(* Logix 5000 project; controller DSFW_Budzar vendor 1 type 14 code 154 rev 32.13; software revision 32.03; part 2 of 5 *)
(* tags used below, declared in another part *)
   ACKNOWLEDGE_ALARMS : BOOL;
   Active_Setpoint : REAL;
   ALARMS : DINT[5];
   ALWAYS_OFF : BOOL;
   Batch_High_High_Temp_Delay : TIMER;
   Batch_High_High_Temp_Setpoint : REAL;
   Batch_Jacket_DT_Temp_Delay : TIMER;
   Batch_Low_Low_Temp_Delay : TIMER;
   Batch_Low_Low_Temp_Setpoint : REAL;
   Batch_Mode_Enable : BOOL;
   C1_Low_Oil_Timer : TIMER;
   C1_MP_Timer : TIMER;
   C1_Run_Proof_Timer : TIMER;
   C_101_AUX : ALIAS FOR Local:1:I.Data.8;
   Comp_Start_Purge_Relay : BOOL;
   Compressor_R404A_Superheat : REAL;
   Condenser_Water_Inlet_Temp_Limit : REAL;
   Condenser_Water_Inlet_Temp_TMR : TIMER;
   CR_002 : ALIAS FOR Local:1:I.Data.0;   // Emergency Stop Safety Relay Status
   CR_01 : ALIAS FOR Local:1:I.Data.15;   // Glycol Tank Low Level Alarm Relay Dry Contact
   CR_108 : ALIAS FOR Local:1:O.Data.0;   // Process Pump Motor Relay (Energizes Contactor M-101)
   CR_109 : ALIAS FOR Local:1:O.Data.5;   // Compressor Motor Relay (Energizes Contactor C-101)
   DCS_Comm_TMR : TIMER;
   DCS_Heartbeat_Returned : DINT;
   DCS_Heartbeat_Returned_Last : DINT;
   EEV_Manual_Relief_Delay : TIMER;   // Oil Management, Delay until Flush begins
   EEV_Manual_Relief_Timer : TIMER;   // Oil Management, Duration of Flush
   FIC_101_Run_PID : BOOL;
   HMI_Batch_Hi_Hi_Temp_Delay : DINT;
   HMI_Batch_Jacket_DT_Temp_Delay : DINT;
   HMI_Batch_Low_Low_Temp_Delay : DINT;
   HMI_Condenser_Water_Inlet_Temp_Delay : DINT;
   HMI_EEV_Manual_Relief_Delay : REAL;   // Oil Management, Delay to start relief entered in minutes.
   HMI_EEV_Manual_Relief_Timer : REAL;   // Oil Management, Relief Duration entered in seconds
   HMI_Jacket_Hi_Hi_Temp_Delay : DINT;
   HMI_Jacket_Hi_Temp_Delay : REAL;
   HMI_Jacket_Low_Low_Temp_Delay : DINT;
   HMI_Jacket_Low_Temp_Delay : REAL;
   HMI_Low_Pump_Suction_Pressure_Delay : REAL;
   HMI_PCV_101_Flush_Time : DINT;
   HMI_R507A_High_Superheat_Timer : DINT;
   HMI_R507A_Low_Pressure_Delay : DINT;
   HMI_R507A_Low_Superheat_Timer : DINT;
   HMI_Remote_State_1 : BOOL;
   HMI_Remote_State_2 : BOOL;
   HMI_Return_Trend_Limits : REAL[2];
   HMI_SP_Trend_Limits : REAL[2];
   HMI_Supply_Trend_Limits : REAL[2];
   HMI_Trend_Data : REAL[3];
   HMI_Valve_Flush_SP : REAL;
   Jacket_Batch_Delta_T : REAL;
   Jacket_Batch_High_Delta_T_Setpoint : REAL;
   Jacket_High_High_Temp_Delay : TIMER;
   Jacket_High_High_Temp_Setpoint : REAL;
   Jacket_High_Temp_Delay : TIMER;
   Jacket_High_Temp_Setpoint : REAL;
   Jacket_Low_Low_Temp_Delay : TIMER;
   Jacket_Low_Low_Temp_Setpoint : REAL;
   Jacket_Low_Temp_Delay : TIMER;
   Jacket_Low_Temp_Setpoint : REAL;
   Low_Pump_Suction_Pressure_Delay : TIMER;
   Low_Pump_Suction_Pressure_Setpoint : REAL;
   M_101_AUX : ALIAS FOR Local:1:I.Data.3;
   Oil_Purge_Fail : BOOL;   // Oil Management, This coil will energize after configured purge retries fail
   Oil_Purge_Retires_Enable : BOOL;
   OMB_101 : ALIAS FOR Local:1:I.Data.12;
   PCV_101_Flush_Timer : TIMER;   // PCV-101 Condenser Hot Water Flush Timer
   PM_101 : ALIAS FOR Local:1:I.Data.1;
   PM_101_StartupTMR : TIMER;   // PM-101 Phase Monitor Startup Delay Alarm Timer
   Process_Pump_Diff_Pressure : REAL;
   PT_101 : BL_Analog_Input;   // Process Supply Pressure
   PT_102 : BL_Analog_Input;   // R404A Compressor Suction Pressure
   PT_103 : BL_Analog_Input;   // R404A Compressor Discharge Pressure
   PT_105 : BL_Analog_Input;   // Condenser Chilled Glycol Return Pressure
   PT_107 : BL_Analog_Input;   // Process Pump Suction Pressure
   Pump_1_Low_Press_Delay : TIMER;
   Pump_High_Pressure_Alarm_Setpoint : REAL;
   Pump_Low_Pressure_Alarm_Setpoint : REAL;
   Pump_RP_ALM_TMR : TIMER;
   R404A_High_Pressure_Setpoint : REAL;
   R404A_High_SH_Setpoint : REAL;
   R404A_High_Superheat_Timer : TIMER;
   R404A_Low_Pressure_Delay : TIMER;
   R404A_Low_Pressure_Setpoint : REAL;
   R404A_Low_SH_Setpoint : REAL;
   R404A_Low_Superheat_Timer : TIMER;
   Ramp_Soak_Current_HMI : DINT;
   Ramp_Soak_Segments_HMI : DINT;
   Ramp_Soak_Segments_HMI_Set : REAL;
   Remote_System_Start : BOOL;   // Remote Start/Stop 0=Stop 1=Start
   Remote_Temp_Setpoint : REAL;   // Remote Temperature Setpoint
   RX_RMPS : RAMP_SOAK;
   Slot_2_Status : DINT;
   Slot_3_Status : DINT;
   Slot_4_Status : DINT;
   Slot_5_Status : DINT;
   Slot_6_Status : DINT;
   Slot_7_Status : DINT;
   Slot_8_Status : DINT;
   Slot_9_Status : DINT;
   Start_Up_Delay : TIMER;
   System_Mode : BOOL;   // 0 = Local Control 1 = Remote Control
   TE_101 : BL_Analog_Input;   // Process Supply Temperature
   TE_102 : BL_Analog_Input;   // Process Return Temperature
   TE_108 : BL_Analog_Input;   // CONDENSER CHILLED GLYCOL INLET TEMPERATURE SENSOR
   Temperature_Setpoint_Max : REAL;   // Maximum Operating Temperature Setpoint (Deg C)
   Temperature_Setpoint_Min : REAL;   // Minimum Operating Temperature Setpoint (Deg C)
   TSH_101 : ALIAS FOR Local:1:I.Data.4;
   Valve_delay_count : REAL;
   Valve_Flush_SP : REAL;
   VESSEL_TEMPERATURE : BL_Analog_Input;   // End User Reactor Temperature
(* A_MainProgram, continued *)

ROUTINE General_Process_Alarms   (* ladder *)
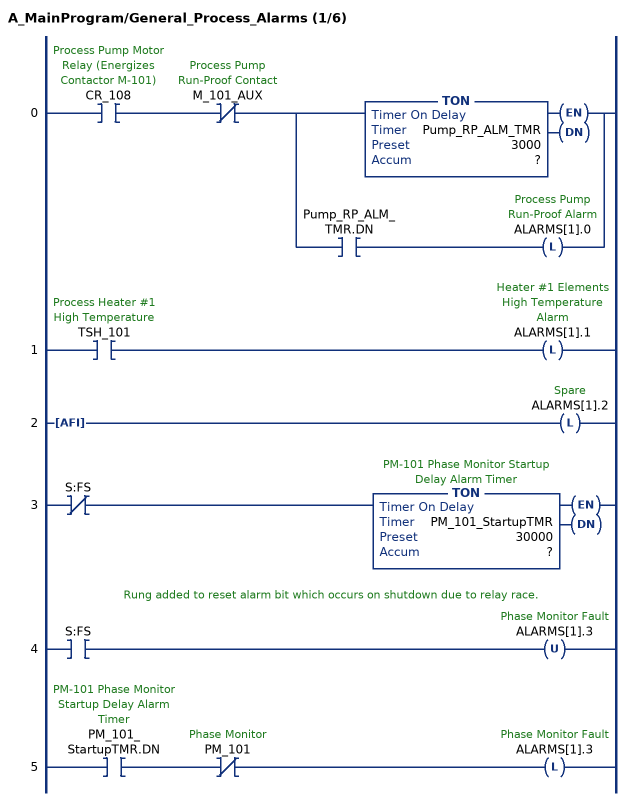
   0: XIC(CR_108)XIO(M_101_AUX)[TON(Pump_RP_ALM_TMR,?,?) ,XIC(Pump_RP_ALM_TMR.DN) OTL(ALARMS[1].0) ];
   1: XIC(TSH_101)OTL(ALARMS[1].1);
   2: AFI()OTL(ALARMS[1].2);
   3: XIO(S:FS)TON(PM_101_StartupTMR,?,?);
   // Rung added to reset alarm bit which occurs on shutdown due to relay race.
   4: XIC(S:FS)OTU(ALARMS[1].3);
   5: XIC(PM_101_StartupTMR.DN)XIO(PM_101)OTL(ALARMS[1].3);
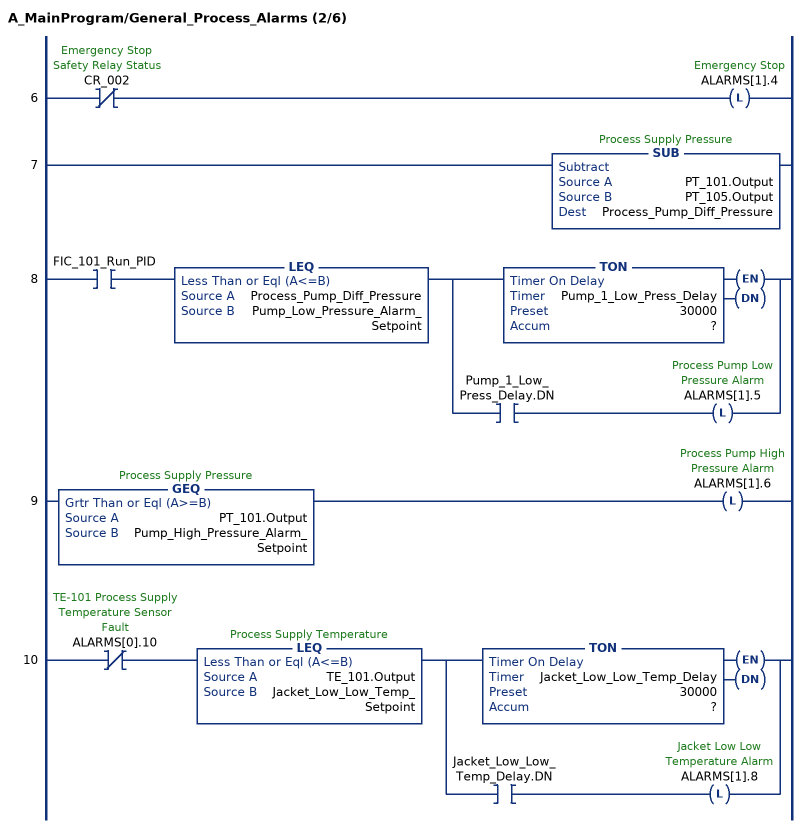
   6: XIO(CR_002)OTL(ALARMS[1].4);
   7: SUB(PT_101.Output,PT_105.Output,Process_Pump_Diff_Pressure);
   8: XIC(FIC_101_Run_PID)LEQ(Process_Pump_Diff_Pressure,Pump_Low_Pressure_Alarm_Setpoint)[TON(Pump_1_Low_Press_Delay,?,?) ,XIC(Pump_1_Low_Press_Delay.DN) OTL(ALARMS[1].5) ];
   9: GEQ(PT_101.Output,Pump_High_Pressure_Alarm_Setpoint)OTL(ALARMS[1].6);
   10: XIO(ALARMS[0].10)LEQ(TE_101.Output,Jacket_Low_Low_Temp_Setpoint)[TON(Jacket_Low_Low_Temp_Delay,?,?) ,XIC(Jacket_Low_Low_Temp_Delay.DN) OTL(ALARMS[1].8) ];
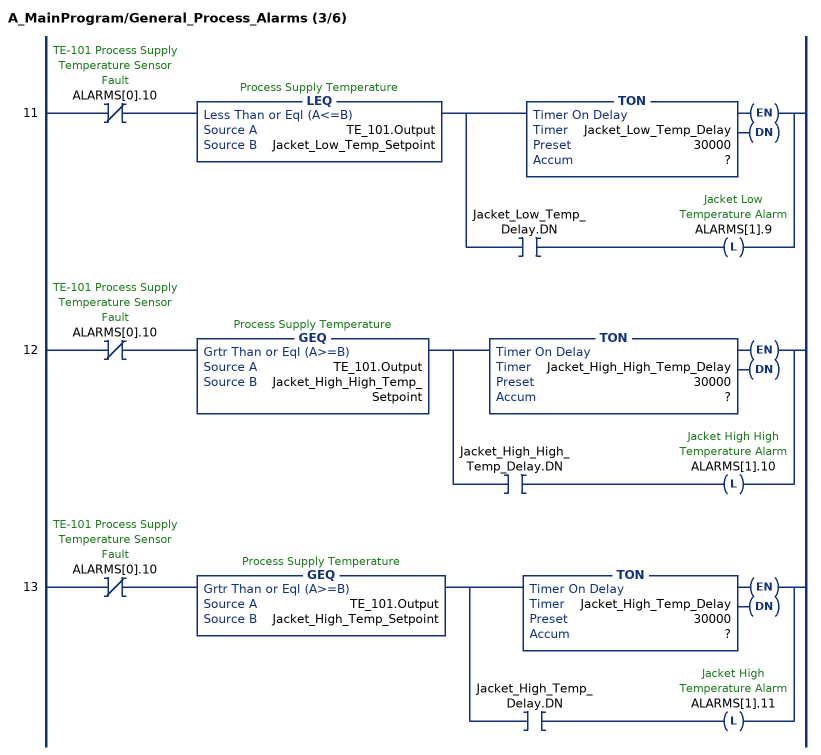
   11: XIO(ALARMS[0].10)LEQ(TE_101.Output,Jacket_Low_Temp_Setpoint)[TON(Jacket_Low_Temp_Delay,?,?) ,XIC(Jacket_Low_Temp_Delay.DN) OTL(ALARMS[1].9) ];
   12: XIO(ALARMS[0].10)GEQ(TE_101.Output,Jacket_High_High_Temp_Setpoint)[TON(Jacket_High_High_Temp_Delay,?,?) ,XIC(Jacket_High_High_Temp_Delay.DN) OTL(ALARMS[1].10) ];
   13: XIO(ALARMS[0].10)GEQ(TE_101.Output,Jacket_High_Temp_Setpoint)[TON(Jacket_High_Temp_Delay,?,?) ,XIC(Jacket_High_Temp_Delay.DN) OTL(ALARMS[1].11) ];
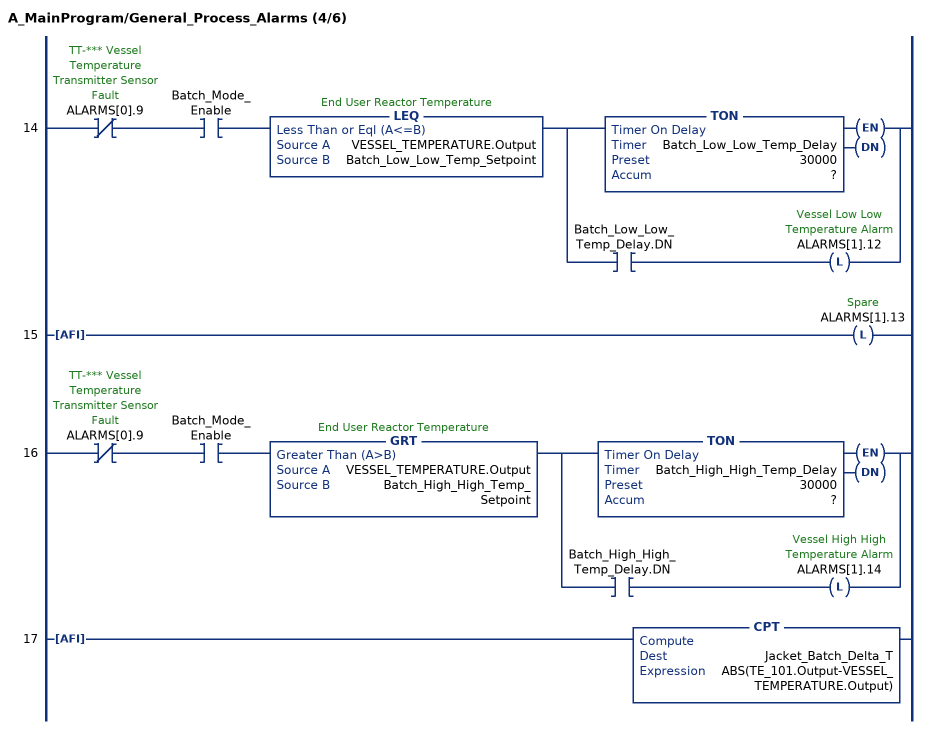
   14: XIO(ALARMS[0].9)XIC(Batch_Mode_Enable)LEQ(VESSEL_TEMPERATURE.Output,Batch_Low_Low_Temp_Setpoint)[TON(Batch_Low_Low_Temp_Delay,?,?) ,XIC(Batch_Low_Low_Temp_Delay.DN) OTL(ALARMS[1].12) ];
   15: AFI()OTL(ALARMS[1].13);
   16: XIO(ALARMS[0].9)XIC(Batch_Mode_Enable)GRT(VESSEL_TEMPERATURE.Output,Batch_High_High_Temp_Setpoint)[TON(Batch_High_High_Temp_Delay,?,?) ,XIC(Batch_High_High_Temp_Delay.DN) OTL(ALARMS[1].14) ];
   17: AFI()CPT(Jacket_Batch_Delta_T,ABS(TE_101.Output-VESSEL_TEMPERATURE.Output));
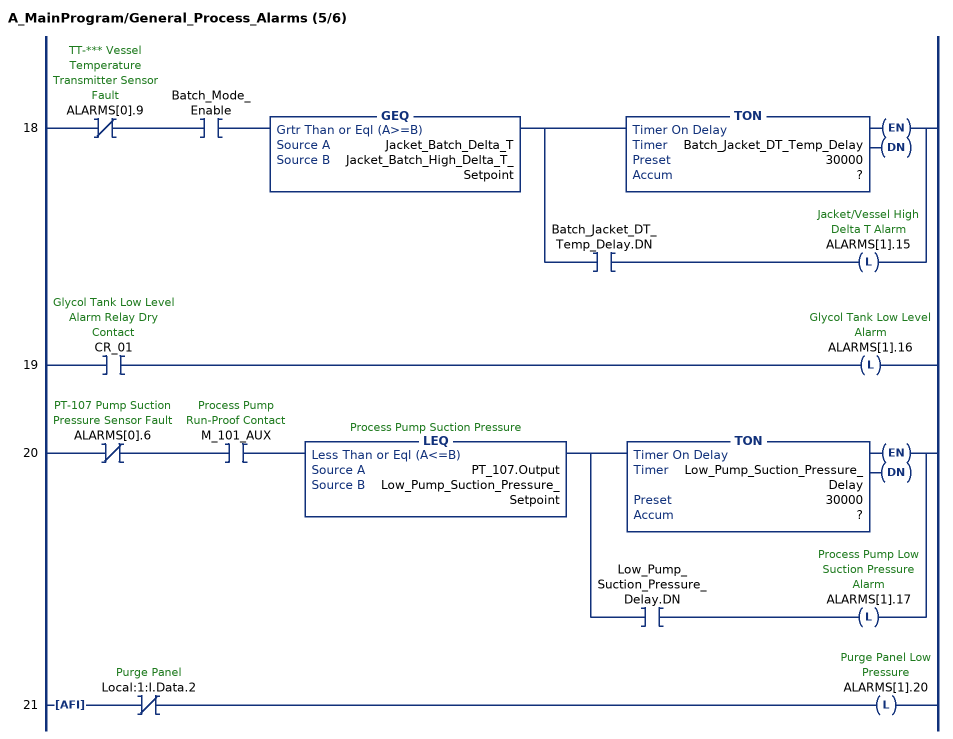
   18: XIO(ALARMS[0].9)XIC(Batch_Mode_Enable)GEQ(Jacket_Batch_Delta_T,Jacket_Batch_High_Delta_T_Setpoint)[TON(Batch_Jacket_DT_Temp_Delay,?,?) ,XIC(Batch_Jacket_DT_Temp_Delay.DN) OTL(ALARMS[1].15) ];
   19: XIC(CR_01)OTL(ALARMS[1].16);
   20: XIO(ALARMS[0].6)XIC(M_101_AUX)LEQ(PT_107.Output,Low_Pump_Suction_Pressure_Setpoint)[TON(Low_Pump_Suction_Pressure_Delay,?,?) ,XIC(Low_Pump_Suction_Pressure_Delay.DN) OTL(ALARMS[1].17) ];
   21: AFI()XIO(Local:1:I.Data.2)OTL(ALARMS[1].20);
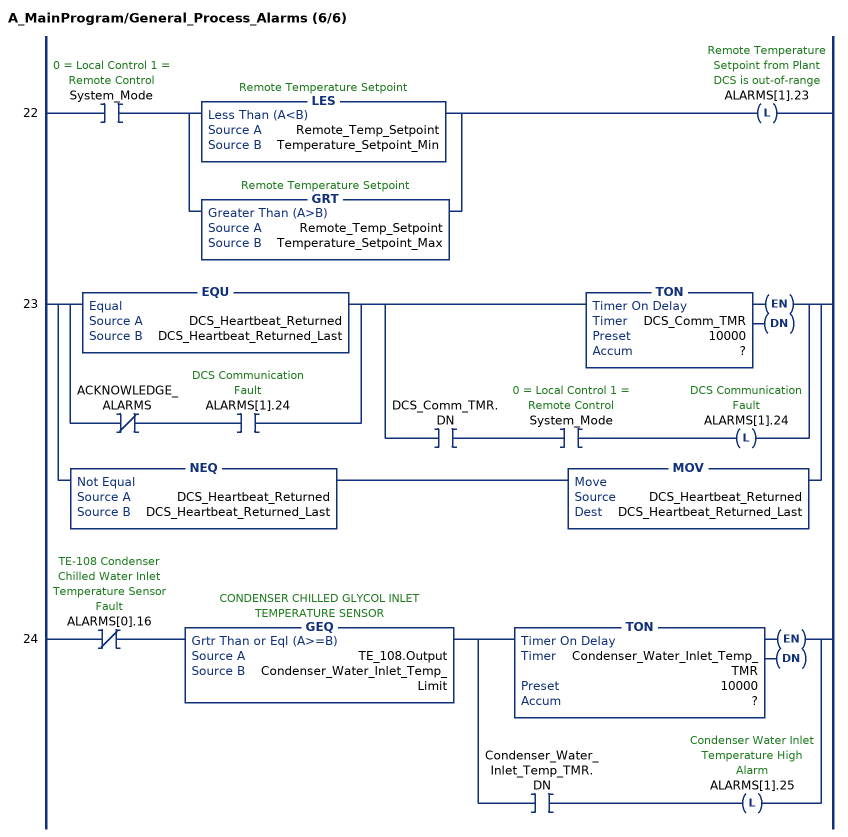
   22: XIC(System_Mode)[LES(Remote_Temp_Setpoint,Temperature_Setpoint_Min) ,GRT(Remote_Temp_Setpoint,Temperature_Setpoint_Max) ]OTL(ALARMS[1].23);
   23: [[EQU(DCS_Heartbeat_Returned,DCS_Heartbeat_Returned_Last) ,XIO(ACKNOWLEDGE_ALARMS) XIC(ALARMS[1].24) ] [TON(DCS_Comm_TMR,?,?) ,XIC(DCS_Comm_TMR.DN) XIC(System_Mode) OTL(ALARMS[1].24) ] ,NEQ(DCS_Heartbeat_Returned,DCS_Heartbeat_Returned_Last) MOV(DCS_Heartbeat_Returned,DCS_Heartbeat_Returned_Last) ];
   24: XIO(ALARMS[0].16)GEQ(TE_108.Output,Condenser_Water_Inlet_Temp_Limit)[TON(Condenser_Water_Inlet_Temp_TMR,?,?) ,XIC(Condenser_Water_Inlet_Temp_TMR.DN) OTL(ALARMS[1].25) ];
END_ROUTINE

ROUTINE HMI_Writes   (* ladder *)
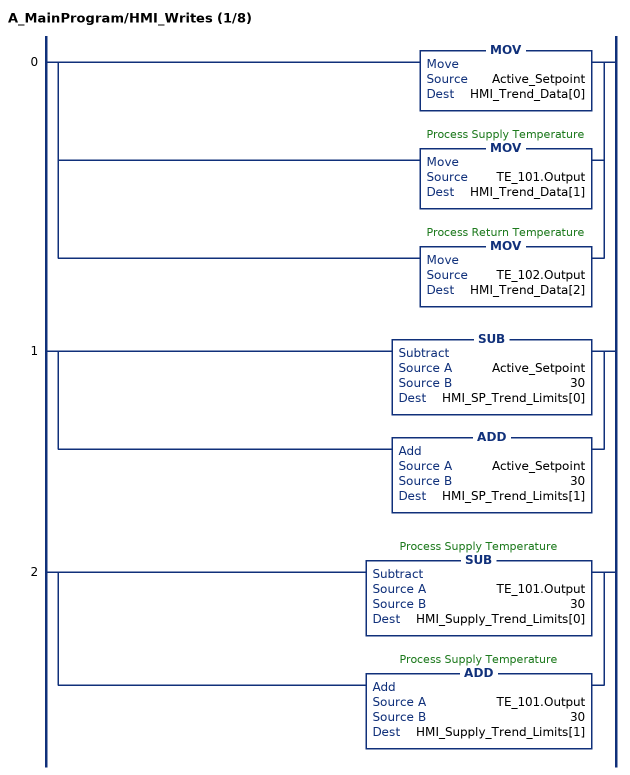
   0: [MOV(Active_Setpoint,HMI_Trend_Data[0]) ,MOV(TE_101.Output,HMI_Trend_Data[1]) ,MOV(TE_102.Output,HMI_Trend_Data[2]) ];
   1: [SUB(Active_Setpoint,30,HMI_SP_Trend_Limits[0]) ,ADD(Active_Setpoint,30,HMI_SP_Trend_Limits[1]) ];
   2: [SUB(TE_101.Output,30,HMI_Supply_Trend_Limits[0]) ,ADD(TE_101.Output,30,HMI_Supply_Trend_Limits[1]) ];
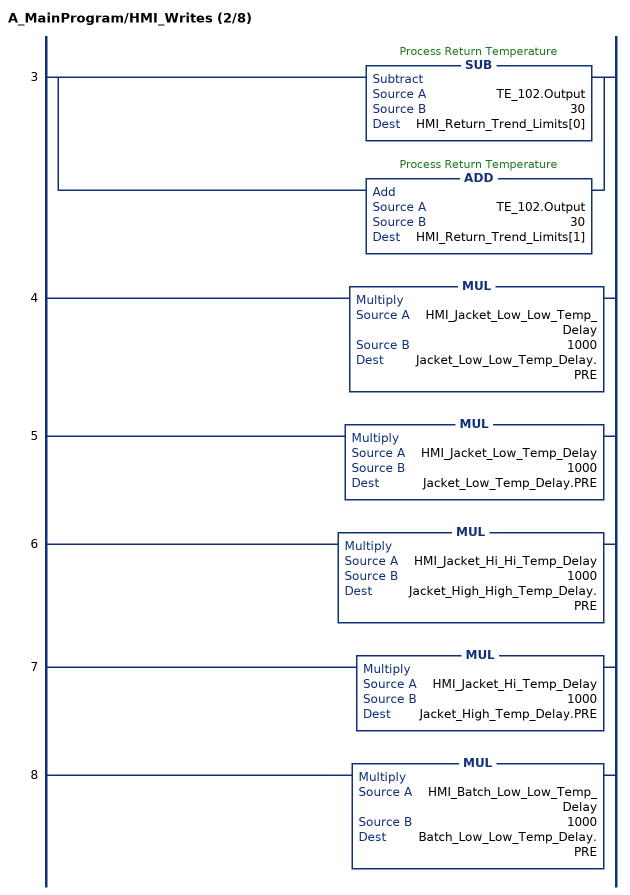
   3: [SUB(TE_102.Output,30,HMI_Return_Trend_Limits[0]) ,ADD(TE_102.Output,30,HMI_Return_Trend_Limits[1]) ];
   4: MUL(HMI_Jacket_Low_Low_Temp_Delay,1000,Jacket_Low_Low_Temp_Delay.PRE);
   5: MUL(HMI_Jacket_Low_Temp_Delay,1000,Jacket_Low_Temp_Delay.PRE);
   6: MUL(HMI_Jacket_Hi_Hi_Temp_Delay,1000,Jacket_High_High_Temp_Delay.PRE);
   7: MUL(HMI_Jacket_Hi_Temp_Delay,1000,Jacket_High_Temp_Delay.PRE);
   8: MUL(HMI_Batch_Low_Low_Temp_Delay,1000,Batch_Low_Low_Temp_Delay.PRE);
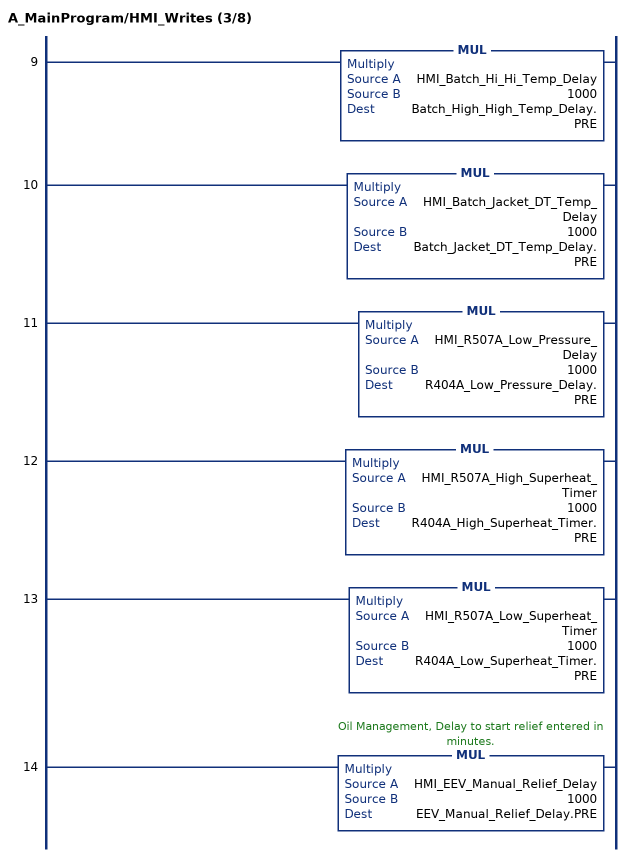
   9: MUL(HMI_Batch_Hi_Hi_Temp_Delay,1000,Batch_High_High_Temp_Delay.PRE);
   10: MUL(HMI_Batch_Jacket_DT_Temp_Delay,1000,Batch_Jacket_DT_Temp_Delay.PRE);
   11: MUL(HMI_R507A_Low_Pressure_Delay,1000,R404A_Low_Pressure_Delay.PRE);
   12: MUL(HMI_R507A_High_Superheat_Timer,1000,R404A_High_Superheat_Timer.PRE);
   13: MUL(HMI_R507A_Low_Superheat_Timer,1000,R404A_Low_Superheat_Timer.PRE);
   14: MUL(HMI_EEV_Manual_Relief_Delay,1000,EEV_Manual_Relief_Delay.PRE);
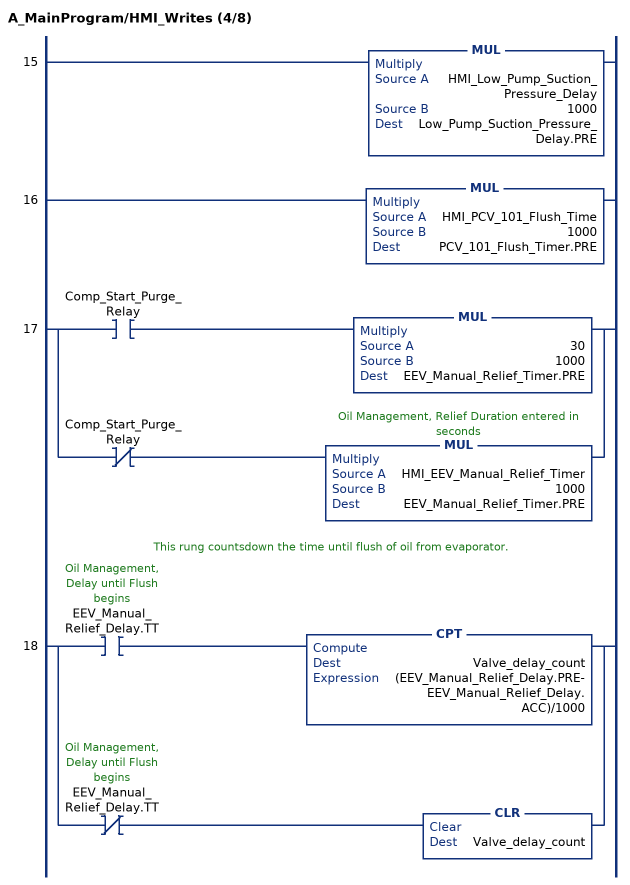
   15: MUL(HMI_Low_Pump_Suction_Pressure_Delay,1000,Low_Pump_Suction_Pressure_Delay.PRE);
   16: MUL(HMI_PCV_101_Flush_Time,1000,PCV_101_Flush_Timer.PRE);
   17: [XIC(Comp_Start_Purge_Relay) MUL(30,1000,EEV_Manual_Relief_Timer.PRE) ,XIO(Comp_Start_Purge_Relay) MUL(HMI_EEV_Manual_Relief_Timer,1000,EEV_Manual_Relief_Timer.PRE) ];
   // This rung countsdown the time until flush of oil from evaporator.
   18: [XIC(EEV_Manual_Relief_Delay.TT) CPT(Valve_delay_count,(EEV_Manual_Relief_Delay.PRE-EEV_Manual_Relief_Delay.ACC)/1000) ,XIO(EEV_Manual_Relief_Delay.TT) CLR(Valve_delay_count) ];
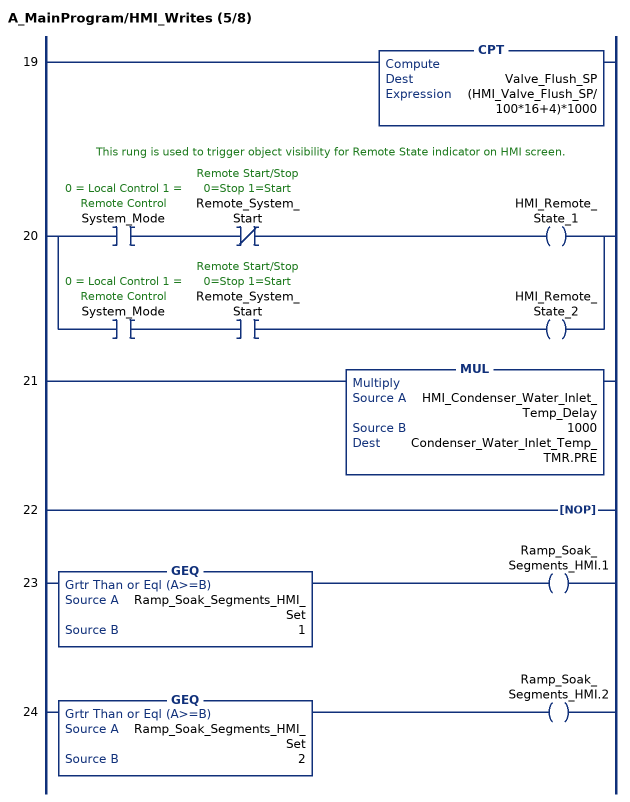
   19: CPT(Valve_Flush_SP,(HMI_Valve_Flush_SP/100*16+4)*1000);
   // This rung is used to trigger object visibility for Remote State indicator on HMI screen.
   20: [XIC(System_Mode) XIO(Remote_System_Start) OTE(HMI_Remote_State_1) ,XIC(System_Mode) XIC(Remote_System_Start) OTE(HMI_Remote_State_2) ];
   21: MUL(HMI_Condenser_Water_Inlet_Temp_Delay,1000,Condenser_Water_Inlet_Temp_TMR.PRE);
   22: NOP();
   23: GEQ(Ramp_Soak_Segments_HMI_Set,1)OTE(Ramp_Soak_Segments_HMI.1);
   24: GEQ(Ramp_Soak_Segments_HMI_Set,2)OTE(Ramp_Soak_Segments_HMI.2);
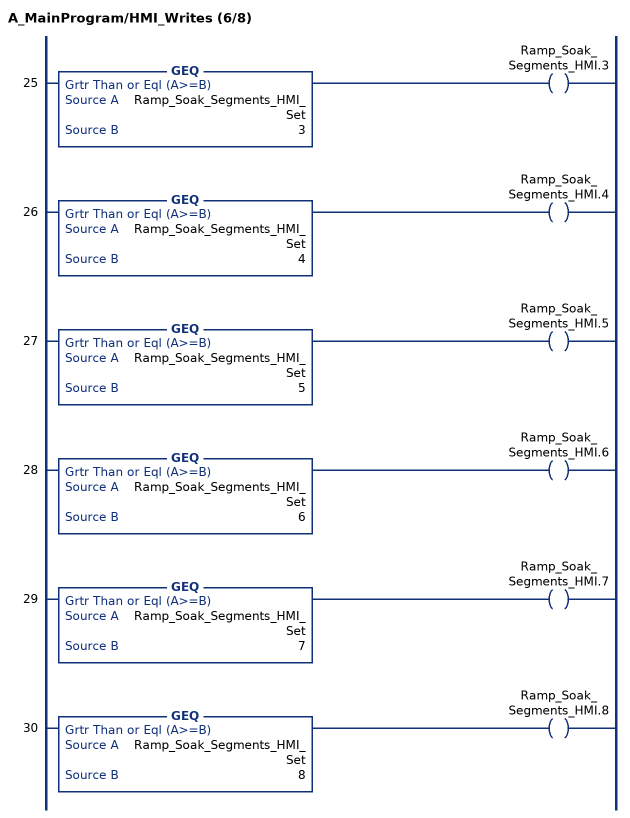
   25: GEQ(Ramp_Soak_Segments_HMI_Set,3)OTE(Ramp_Soak_Segments_HMI.3);
   26: GEQ(Ramp_Soak_Segments_HMI_Set,4)OTE(Ramp_Soak_Segments_HMI.4);
   27: GEQ(Ramp_Soak_Segments_HMI_Set,5)OTE(Ramp_Soak_Segments_HMI.5);
   28: GEQ(Ramp_Soak_Segments_HMI_Set,6)OTE(Ramp_Soak_Segments_HMI.6);
   29: GEQ(Ramp_Soak_Segments_HMI_Set,7)OTE(Ramp_Soak_Segments_HMI.7);
   30: GEQ(Ramp_Soak_Segments_HMI_Set,8)OTE(Ramp_Soak_Segments_HMI.8);
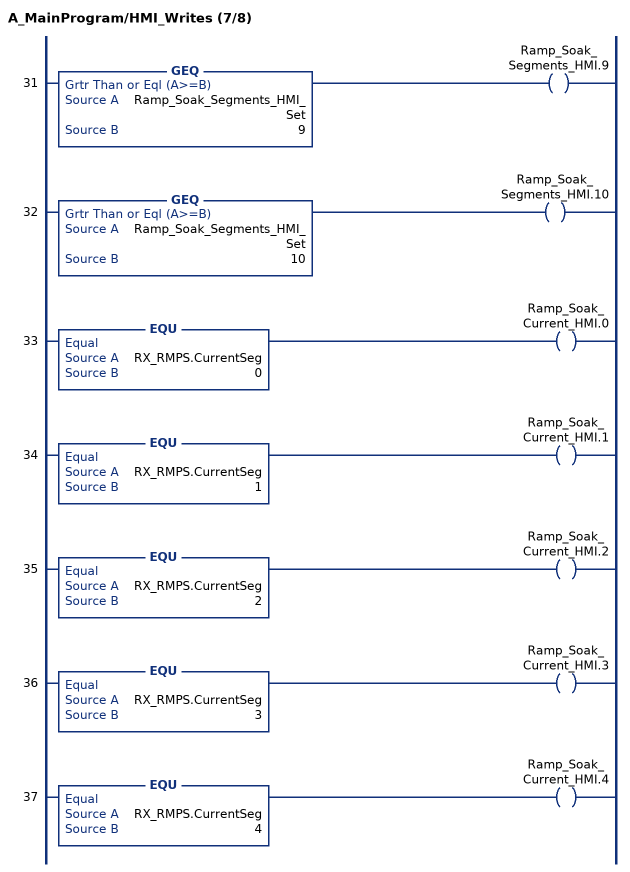
   31: GEQ(Ramp_Soak_Segments_HMI_Set,9)OTE(Ramp_Soak_Segments_HMI.9);
   32: GEQ(Ramp_Soak_Segments_HMI_Set,10)OTE(Ramp_Soak_Segments_HMI.10);
   33: EQU(RX_RMPS.CurrentSeg,0)OTE(Ramp_Soak_Current_HMI.0);
   34: EQU(RX_RMPS.CurrentSeg,1)OTE(Ramp_Soak_Current_HMI.1);
   35: EQU(RX_RMPS.CurrentSeg,2)OTE(Ramp_Soak_Current_HMI.2);
   36: EQU(RX_RMPS.CurrentSeg,3)OTE(Ramp_Soak_Current_HMI.3);
   37: EQU(RX_RMPS.CurrentSeg,4)OTE(Ramp_Soak_Current_HMI.4);
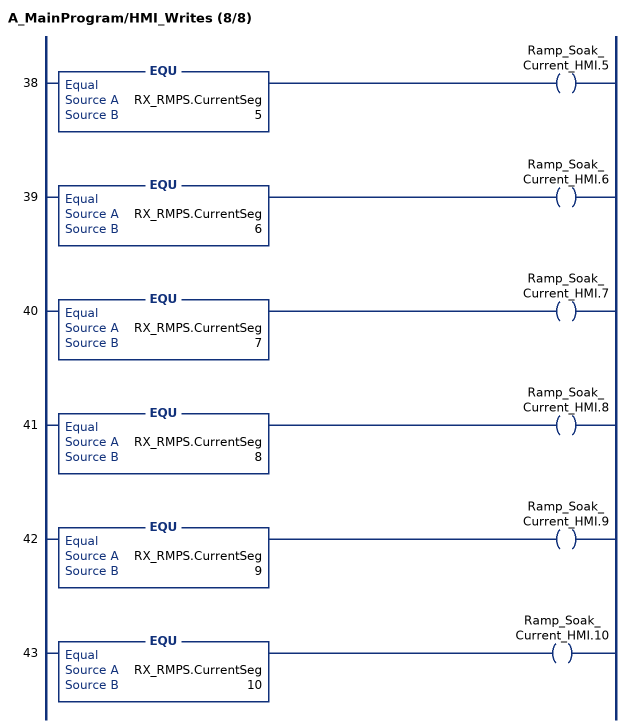
   38: EQU(RX_RMPS.CurrentSeg,5)OTE(Ramp_Soak_Current_HMI.5);
   39: EQU(RX_RMPS.CurrentSeg,6)OTE(Ramp_Soak_Current_HMI.6);
   40: EQU(RX_RMPS.CurrentSeg,7)OTE(Ramp_Soak_Current_HMI.7);
   41: EQU(RX_RMPS.CurrentSeg,8)OTE(Ramp_Soak_Current_HMI.8);
   42: EQU(RX_RMPS.CurrentSeg,9)OTE(Ramp_Soak_Current_HMI.9);
   43: EQU(RX_RMPS.CurrentSeg,10)OTE(Ramp_Soak_Current_HMI.10);
END_ROUTINE

ROUTINE IO_Module_Fault   (* ladder *)
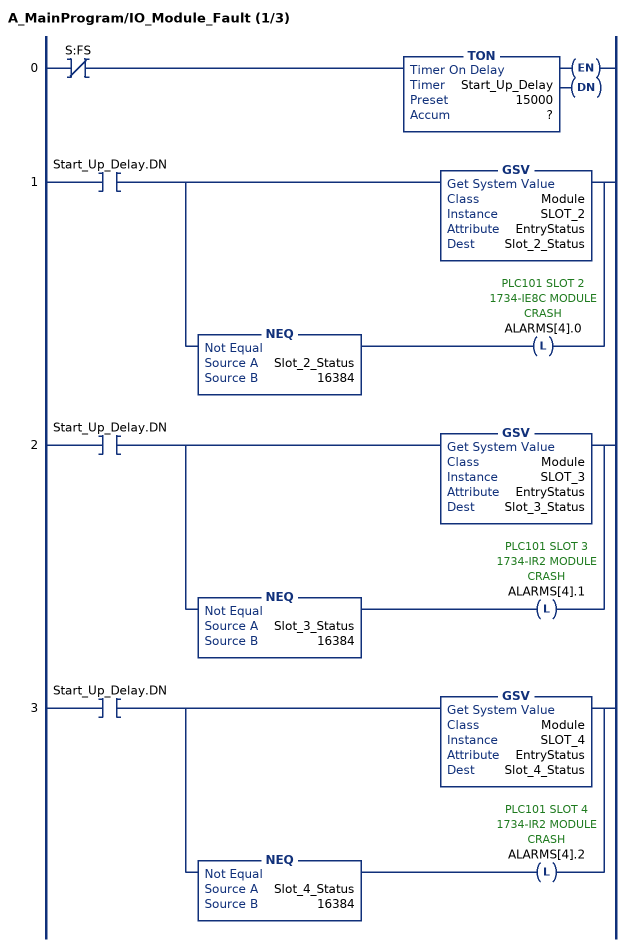
   0: XIO(S:FS)TON(Start_Up_Delay,?,?);
   1: XIC(Start_Up_Delay.DN)[GSV(Module,SLOT_2,EntryStatus,Slot_2_Status) ,NEQ(Slot_2_Status,16384) OTL(ALARMS[4].0) ];
   2: XIC(Start_Up_Delay.DN)[GSV(Module,SLOT_3,EntryStatus,Slot_3_Status) ,NEQ(Slot_3_Status,16384) OTL(ALARMS[4].1) ];
   3: XIC(Start_Up_Delay.DN)[GSV(Module,SLOT_4,EntryStatus,Slot_4_Status) ,NEQ(Slot_4_Status,16384) OTL(ALARMS[4].2) ];
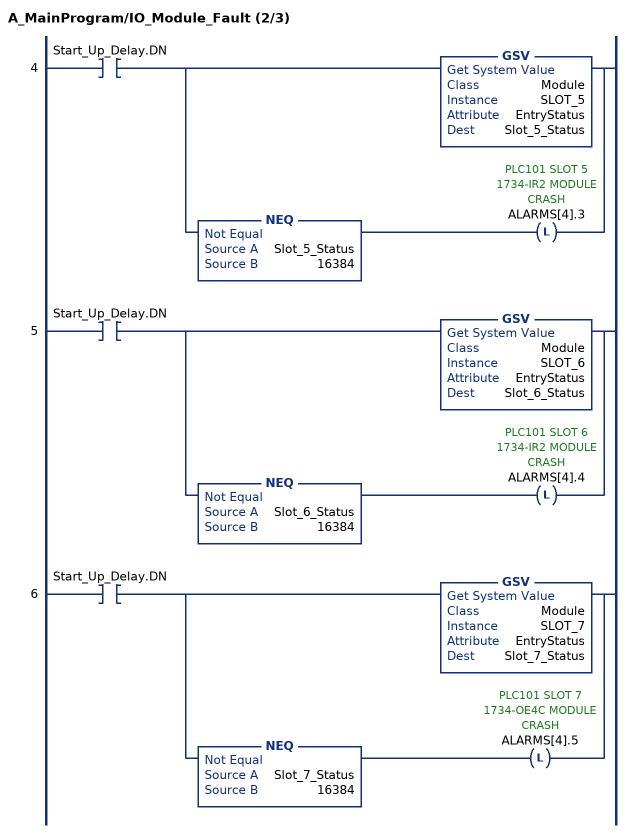
   4: XIC(Start_Up_Delay.DN)[GSV(Module,SLOT_5,EntryStatus,Slot_5_Status) ,NEQ(Slot_5_Status,16384) OTL(ALARMS[4].3) ];
   5: XIC(Start_Up_Delay.DN)[GSV(Module,SLOT_6,EntryStatus,Slot_6_Status) ,NEQ(Slot_6_Status,16384) OTL(ALARMS[4].4) ];
   6: XIC(Start_Up_Delay.DN)[GSV(Module,SLOT_7,EntryStatus,Slot_7_Status) ,NEQ(Slot_7_Status,16384) OTL(ALARMS[4].5) ];
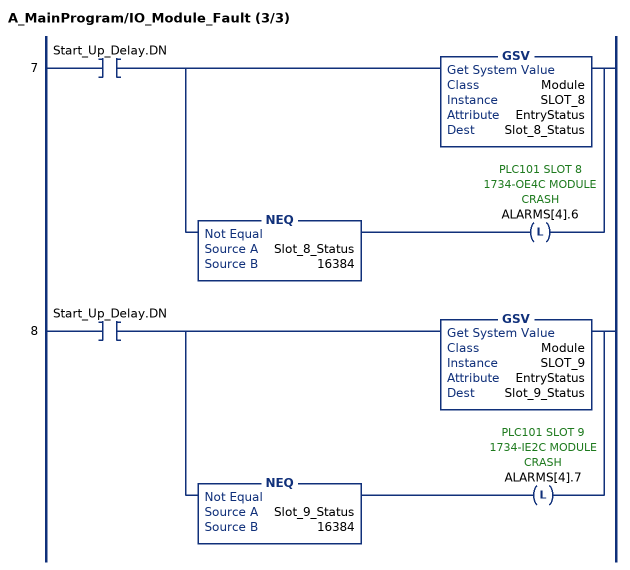
   7: XIC(Start_Up_Delay.DN)[GSV(Module,SLOT_8,EntryStatus,Slot_8_Status) ,NEQ(Slot_8_Status,16384) OTL(ALARMS[4].6) ];
   8: XIC(Start_Up_Delay.DN)[GSV(Module,SLOT_9,EntryStatus,Slot_9_Status) ,NEQ(Slot_9_Status,16384) OTL(ALARMS[4].7) ];
END_ROUTINE

ROUTINE R404A_Alarms   (* ladder *)
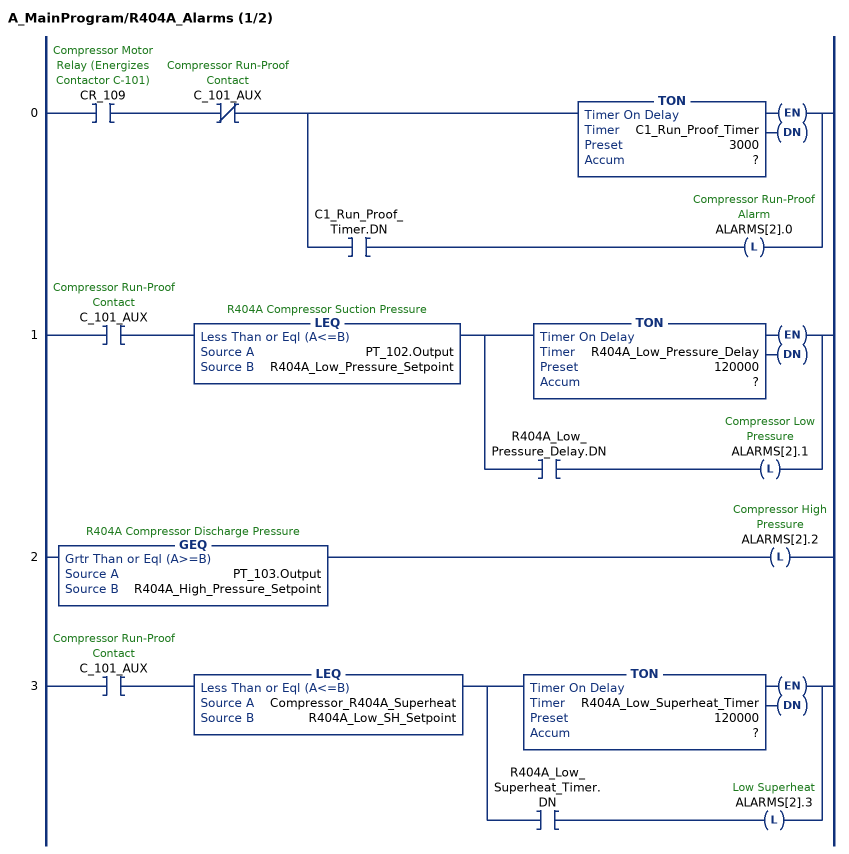
   0: XIC(CR_109)XIO(C_101_AUX)[TON(C1_Run_Proof_Timer,?,?) ,XIC(C1_Run_Proof_Timer.DN) OTL(ALARMS[2].0) ];
   1: XIC(C_101_AUX)LEQ(PT_102.Output,R404A_Low_Pressure_Setpoint)[TON(R404A_Low_Pressure_Delay,?,?) ,XIC(R404A_Low_Pressure_Delay.DN) OTL(ALARMS[2].1) ];
   2: GEQ(PT_103.Output,R404A_High_Pressure_Setpoint)OTL(ALARMS[2].2);
   3: XIC(C_101_AUX)LEQ(Compressor_R404A_Superheat,R404A_Low_SH_Setpoint)[TON(R404A_Low_Superheat_Timer,?,?) ,XIC(R404A_Low_Superheat_Timer.DN) OTL(ALARMS[2].3) ];
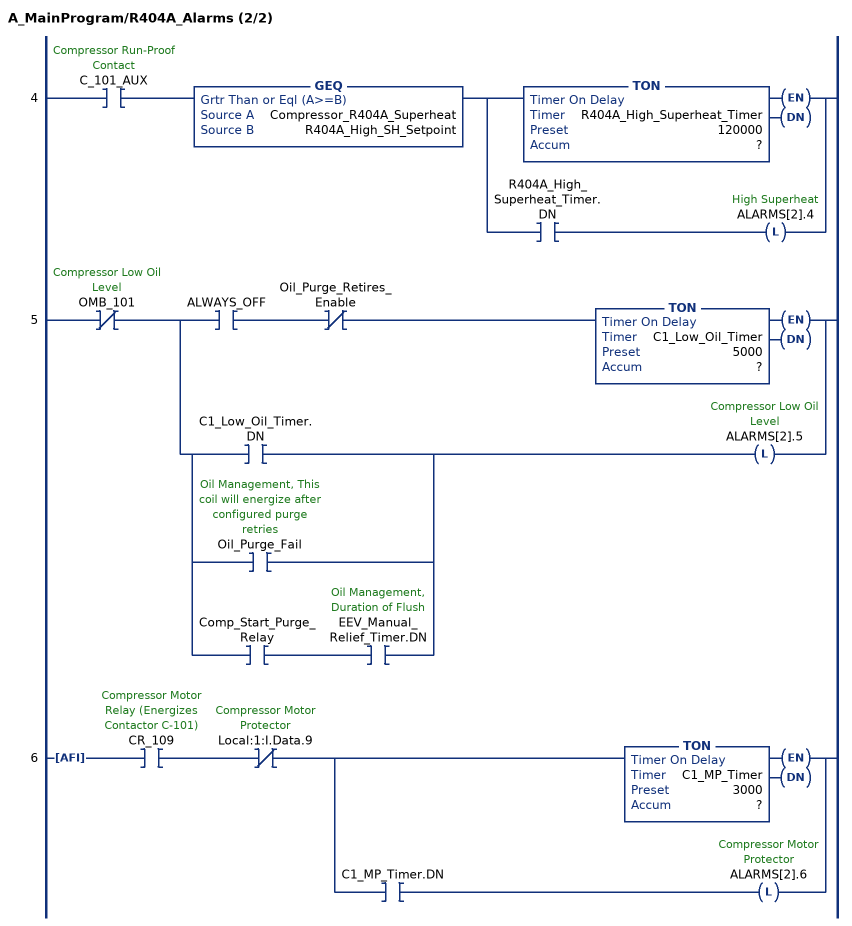
   4: XIC(C_101_AUX)GEQ(Compressor_R404A_Superheat,R404A_High_SH_Setpoint)[TON(R404A_High_Superheat_Timer,?,?) ,XIC(R404A_High_Superheat_Timer.DN) OTL(ALARMS[2].4) ];
   5: XIO(OMB_101)[XIC(ALWAYS_OFF) XIO(Oil_Purge_Retires_Enable) TON(C1_Low_Oil_Timer,?,?) ,[XIC(C1_Low_Oil_Timer.DN) ,XIC(Oil_Purge_Fail) ,XIC(Comp_Start_Purge_Relay) XIC(EEV_Manual_Relief_Timer.DN) ] OTL(ALARMS[2].5) ];
   6: AFI()XIC(CR_109)XIO(Local:1:I.Data.9)[TON(C1_MP_Timer,?,?) ,XIC(C1_MP_Timer.DN) OTL(ALARMS[2].6) ];
END_ROUTINE
